// TIA Portal V21 export
// export: Created 2026-11-10T07:27:30.7974892Z, ExportSetting WithDefaults, DisplayName Totally Integrated Automation Portal, DisplayVersion V21 Update 3, DisplayName STEP 7 Professional, DisplayVersion V21 Update 3, DisplayName STEP 7 Safety, DisplayVersion V21, DisplayName Tech WebApplication, DisplayVersion V21, DisplayName WinCC Basic/Comfort/Advanced, DisplayVersion V21 Update 3, DisplayName WinCC Unified, DisplayVersion V21 Update 3
FUNCTION_BLOCK "FB_LadTech"   // FB5, LAD
{ S7_Optimized_Access := 'TRUE' }
VERSION : 0.1
// stored: AutoNumber true, IsIECCheckEnabled false, IsRetainMemResEnabled false, MemoryReserve 100, SetENOAutomatically false, UDAEnableTagReadback false
   VAR_INPUT
      sp : Real;
      pv : Real;
   END_VAR
   VAR_OUTPUT
      outv : Real;
      err : Bool;
   END_VAR
BEGIN

REGION Network 1: PID call
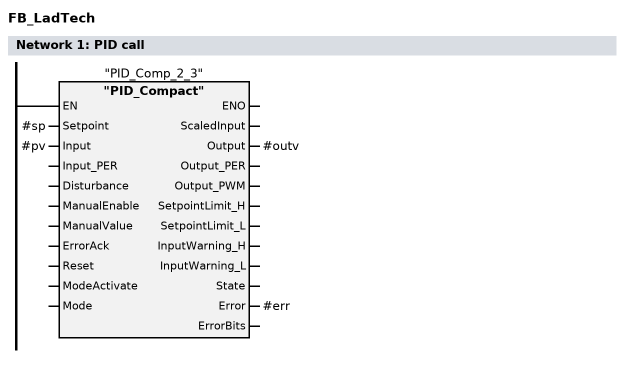
   RUNG wire#powerrail
      "PID_Comp_2_3"(Setpoint := #sp, Input := #pv, Output => #outv, Error => #err, Input_PER :=, Disturbance :=, ManualEnable :=, ManualValue :=, ErrorAck :=, Reset :=, ModeActivate :=, ScaledInput =>, Output_PER =>, Output_PWM =>, SetpointLimit_H =>, SetpointLimit_L =>, InputWarning_H =>, InputWarning_L =>, State =>, ErrorBits =>, Mode :=)
   END_RUNG
   // the same network as SCL:
   "PID_Comp_2_3"(Setpoint := #sp, Input := #pv, Output => #outv, Error => #err);   // "PID_Compact"
END_REGION
END_FUNCTION_BLOCK
